(* IEC 61131-3 sources: CannyIECUnitTest/st/device/plc_logic/application, 3 files *)

(* ---- testcase-TestCase.st ---- *)
(* --- Interface --- *)
{attribute 'test'}
{attribute 'testcasename':='ArrayOfLag'}
{attribute 'testcasetimeout':='15000'}
FUNCTION_BLOCK TestCase EXTENDS TM.Testcase
VAR_INPUT
END_VAR
VAR_OUTPUT
END_VAR
VAR
END_VAR

(* --- Implementation --- *)
SUPER^();

(* ---- testcase_isignbit-TestCase_ISIGNBIT.st ---- *)
(* --- Interface --- *)
{attribute 'test'}
{attribute 'testcasename':='ArrayOfLag'}
{attribute 'testcasetimeout':='15000'}
FUNCTION_BLOCK TestCase_ISIGNBIT EXTENDS Testcase
VAR_INPUT
END_VAR
VAR_OUTPUT
END_VAR
VAR
END_VAR

(* --- Implementation --- *)
SUPER^();

(* ---- plc_prg-PLC_PRG.st ---- *)
(* --- Interface --- *)
PROGRAM PLC_PRG
VAR
	fbTestCase : TestCase_ISIGNBIT;
END_VAR
